// TIA Portal V20 export
Screen "Pop-up_MOVE_LEGEND_Popup"  400x505
  ScreenItem "Rechteck_1" at 0,0 size 400x505  Type=HmiRectangle
  ScreenItem "Textfeld_Legende" at 1,1 size 398x25  Type=HmiTextBox
  ScreenItem "Arrow_ADV_Left_Fast" at 24,195 size 15x30  Type=HmiPolygon
  ScreenItem "Arrow_RTN_Right_Fast" at 78,195 size 15x30  Type=HmiPolygon
  ScreenItem "Textfeld_2" at 10,125 size 165x20  Type=HmiTextBox
  ScreenItem "Textfeld_1" at 10,147 size 165x20  Type=HmiTextBox
  ScreenItem "Textfeld_3" at 10,37 size 165x20  Type=HmiTextBox
  ScreenItem "Textfeld_4" at 10,59 size 165x20  Type=HmiTextBox
  ScreenItem "Textfeld_5" at 10,81 size 165x20  Type=HmiTextBox
  ScreenItem "Textfeld_6" at 10,103 size 165x20  Type=HmiTextBox
  ScreenItem "Textfeld_9" at 180,125 size 165x20  Type=HmiTextBox
  ScreenItem "Textfeld_10" at 180,147 size 165x20  Type=HmiTextBox
  ScreenItem "Textfeld_11" at 180,37 size 120x20  Type=HmiTextBox
  ScreenItem "Textfeld_12" at 180,59 size 200x20  Type=HmiTextBox
  ScreenItem "Textfeld_13" at 180,74 size 141x33  Type=HmiTextBox
  ScreenItem "Textfeld_14" at 180,103 size 165x20  Type=HmiTextBox
  ScreenItem "Textfeld_15" at 10,172 size 100x20  Type=HmiTextBox
  ScreenItem "Textfeld_16" at 109,190 size 280x40  Type=HmiTextBox
  ScreenItem "Textfeld_17" at 109,232 size 280x20  Type=HmiTextBox
  ScreenItem "Textfeld_18" at 109,259 size 280x20  Type=HmiTextBox
  ScreenItem "Cancel Mode" at 309,1 size 90x60  Type=HmiButton
  ScreenItem "PB_ADV" at 13,230 size 36x24  Type=HmiButton
  ScreenItem "PB_RTN" at 67,230 size 36x24  Type=HmiButton
  ScreenItem "PB_ADV_1" at 13,257 size 36x24  Type=HmiButton
  ScreenItem "PB_RTN_1" at 67,257 size 36x24  Type=HmiButton
  ScreenItem "PB_ON" at 13,284 size 36x24  Type=HmiButton
  ScreenItem "PB_OFF" at 67,284 size 36x24  Type=HmiButton
  ScreenItem "Safety" at 13,445 size 90x25  Type=HmiButton
  ScreenItem "Teil_vorh" at 13,416 size 90x25  Type=HmiButton
  ScreenItem "Position_LeftEnd" at 13,311 size 30x20  Type=HmiTextBox
  ScreenItem "Position_LeftSlow" at 73,311 size 30x20  Type=HmiTextBox
  ScreenItem "InterlockADV" at 13,389 size 90x25  Type=HmiButton
  ScreenItem "ADV_Fast" at 13,361 size 90x25  Type=HmiButton
  ScreenItem "ADV_Slow" at 13,334 size 90x25  Type=HmiButton
  ScreenItem "Feedback DeviceON" at 13,473 size 90x25  Type=HmiButton
  ScreenItem "Textfeld_7" at 109,286 size 280x20  Type=HmiTextBox
  ScreenItem "Textfeld_8" at 109,309 size 280x20  Type=HmiTextBox
  ScreenItem "Textfeld_19" at 109,335 size 280x20  Type=HmiTextBox
  ScreenItem "Textfeld_20" at 109,363 size 280x20  Type=HmiTextBox
  ScreenItem "Textfeld_21" at 109,390 size 280x20  Type=HmiTextBox
  ScreenItem "Textfeld_22" at 109,418 size 280x20  Type=HmiTextBox
  ScreenItem "Textfeld_23" at 109,446 size 280x20  Type=HmiTextBox
  ScreenItem "Textfeld_24" at 109,476 size 280x20  Type=HmiTextBox
